(* IEC 61131-3 sources: NachHouse_TST/API/pilot_API_V10, 4 files *)

(* ---- 01_Nh_Api_STRUCT.st ---- *)
// NachHouse API PLC pilot V1.
// The public contract uses native PLCComS PUBLIC_API variables only.
// SK: Verejny kontrakt pouziva iba nativne PUBLIC_API premenne PLCComS.

VAR_GLOBAL CONSTANT
   NH_API_PROTOCOL_VERSION       : UINT := 1;            // Binary protocol version. SK: Verzia binarneho protokolu.
   NH_API_MAGIC                  : DWORD := 16#5041484E;  // ASCII NHAP bytes in little-endian order. SK: Bajty ASCII NHAP v little-endian poradi.
   NH_API_HEADER_SIZE            : UINT := 64;           // Fixed header size in bytes. SK: Pevna velkost hlavicky v bajtoch.
   NH_API_TX_WORD_COUNT          : UINT := 512;          // Number of DWORD words in the shared TX buffer. SK: Pocet DWORD slov spolocneho TX buffera.
   NH_API_RX_WORDS_PER_CLIENT    : UINT := 64;           // DWORD words in one client RX segment. SK: Pocet DWORD slov RX segmentu jedneho klienta.
   NH_API_RX_WORD_COUNT          : UINT := 256;          // Four RX segments of 64 DWORD each. SK: Styri RX segmenty po 64 DWORD.
   NH_API_MAX_CLIENTS            : USINT := 4;           // Maximum concurrently registered clients. SK: Najvacsi pocet sucasne registrovanych klientov.
   NH_API_MAX_ROOMS              : USINT := 40;          // Maximum number of pilot rooms. SK: Najvacsi pocet miestnosti pilotu.

   NH_API_CONFIG_RECORD_SIZE     : UINT := 138;          // Wire config record size. SK: Velkost wire config zaznamu.
   NH_API_STATE_RECORD_SIZE      : UINT := 22;           // Wire state record size including Twilight. SK: Velkost wire state zaznamu vratane Twilight.
   NH_API_CONFIG_DIFF_SIZE       : UINT := 143;          // Operation, RoomId and config record. SK: Operacia, RoomId a config zaznam.
   NH_API_STATE_DIFF_SIZE        : UINT := 27;           // Operation, RoomId and state record. SK: Operacia, RoomId a state zaznam.
   NH_API_CONFIG_PER_FRAME       : USINT := 14;          // Maximum config records in one TX frame. SK: Najviac config zaznamov v jednom TX ramci.
   NH_API_STATE_PER_FRAME        : USINT := 40;          // Maximum state records in one TX frame. SK: Najviac state zaznamov v jednom TX ramci.
   NH_API_CONFIG_DIFF_PER_FRAME  : USINT := 13;          // Maximum config changes in one TX frame. SK: Najviac config zmien v jednom TX ramci.
   NH_API_STATE_DIFF_PER_FRAME   : USINT := 40;          // Maximum state changes in one TX frame. SK: Najviac state zmien v jednom TX ramci.

   NH_API_TX_IDLE                : USINT := 0;            // TX buffer may be built. SK: TX buffer sa moze naplnit.
   NH_API_TX_BUILDING            : USINT := 1;            // PLC is building a TX frame. SK: PLC prave pripravuje TX ramec.
   NH_API_TX_READY               : USINT := 2;            // TX frame is stable and waiting for ACK. SK: TX ramec je stabilny a caka na ACK.

   NH_API_CLIENT_FREE            : USINT := 0;            // Client slot is free. SK: Klientsky slot je volny.
   NH_API_CLIENT_ACTIVE          : USINT := 1;            // Client slot has a valid lease. SK: Klientsky slot ma platny lease.

   NH_API_MSG_SNAPSHOT_REQUEST   : UINT := 1;             // RX full snapshot request. SK: RX poziadavka na kompletny snapshot.
   NH_API_MSG_ADD_ROOM           : UINT := 2;             // RX add-room request. SK: RX poziadavka na pridanie miestnosti.
   NH_API_MSG_DELETE_ROOM        : UINT := 3;             // RX delete-room request. SK: RX poziadavka na zmazanie miestnosti.
   NH_API_MSG_COPY_ROOM          : UINT := 4;             // RX copy-room request. SK: RX poziadavka na kopirovanie miestnosti.
   NH_API_MSG_SET_ROOM_CONFIG     : UINT := 5;             // RX room-config update request. SK: RX poziadavka na zmenu configu.
   NH_API_MSG_SET_ROOM_STATE      : UINT := 6;             // RX test room-state update request. SK: RX testovacia poziadavka na zmenu state.
   NH_API_MSG_CONFIG_SNAPSHOT    : UINT := 101;           // TX config snapshot part. SK: TX cast config snapshotu.
   NH_API_MSG_STATE_SNAPSHOT     : UINT := 102;           // TX state snapshot part. SK: TX cast state snapshotu.
   NH_API_MSG_CONFIG_DIFF        : UINT := 103;           // TX config diff. SK: TX config diff.
   NH_API_MSG_STATE_DIFF         : UINT := 104;           // TX state diff. SK: TX state diff.
   NH_API_MSG_SNAPSHOT_DONE      : UINT := 105;           // TX snapshot transaction completion. SK: TX ukoncenie snapshot transakcie.

   NH_API_SCHEMA_NONE            : UINT := 0;             // Message has no data record. SK: Sprava nema datovy zaznam.
   NH_API_SCHEMA_ROOM_CONFIG     : UINT := 1;             // Room configuration schema. SK: Schema konfiguracie miestnosti.
   NH_API_SCHEMA_ROOM_STATE      : UINT := 2;             // Room dynamic-state schema. SK: Schema dynamickeho stavu miestnosti.
   NH_API_SCHEMA_VERSION         : UINT := 1;             // Version of both room schemas. SK: Verzia oboch room schem.

   NH_API_CHANGE_UPSERT          : USINT := 1;            // Insert or complete record update. SK: Pridanie alebo uplna aktualizacia zaznamu.
   NH_API_CHANGE_DELETE          : USINT := 2;            // Record deletion. SK: Odstranenie zaznamu.

   NH_API_RESULT_NONE            : USINT := 0;            // No result is available yet. SK: Vysledok este neexistuje.
   NH_API_RESULT_OK              : USINT := 1;            // Request succeeded. SK: Poziadavka bola uspesna.
   NH_API_RESULT_BUSY            : USINT := 2;            // Another global transaction is active. SK: Ina globalna transakcia este bezi.
   NH_API_RESULT_BAD_FRAME       : USINT := 3;            // Header, size or CRC is invalid. SK: Hlavicka, velkost alebo CRC su neplatne.
   NH_API_RESULT_NOT_FOUND       : USINT := 4;            // Requested room does not exist. SK: Pozadovana miestnost neexistuje.
   NH_API_RESULT_NO_FREE_SLOT    : USINT := 5;            // No room or client slot is free. SK: Nie je volny room alebo client slot.
   NH_API_RESULT_ALREADY_EXISTS  : USINT := 6;            // RoomId already exists. SK: RoomId uz existuje.
   NH_API_RESULT_INVALID         : USINT := 7;            // Request payload is invalid. SK: Obsah poziadavky nie je platny.
   NH_API_RESULT_UNSUPPORTED     : USINT := 8;            // Message type is unsupported. SK: Typ spravy nie je podporovany.

   NH_API_TEST_NONE              : USINT := 0;            // WebMaker performs no action. SK: WebMaker nevykona ziadnu akciu.
   NH_API_TEST_SET_STATE         : USINT := 1;            // WebMaker changes room state. SK: WebMaker zmeni stav miestnosti.
   NH_API_TEST_ADD_ROOM          : USINT := 2;            // WebMaker adds a room. SK: WebMaker prida miestnost.
   NH_API_TEST_DELETE_ROOM       : USINT := 3;            // WebMaker deletes a room. SK: WebMaker zmaze miestnost.
   NH_API_TEST_COPY_ROOM         : USINT := 4;            // WebMaker copies a room. SK: WebMaker skopiruje miestnost.
   NH_API_TEST_SET_CONFIG        : USINT := 5;            // WebMaker changes room config. SK: WebMaker zmeni config miestnosti.
   NH_API_TEST_REQUEST_SNAPSHOT  : USINT := 6;            // WebMaker starts a broadcast snapshot. SK: WebMaker vyvola broadcast snapshot.
END_VAR

TYPE
   NH_ROOM_CONFIG : STRUCT // Static room configuration transferred in snapshots, diffs and commands. SK: Staticka konfiguracia miestnosti prenasana v snapshotoch, diffoch a prikazoch.
      Used           : BOOL;       // TRUE marks an occupied internal slot. SK: TRUE oznacuje obsadeny interny slot.
      RoomId         : UDINT;      // Stable unique room identifier. SK: Stabilny jedinecny identifikator miestnosti.
      Name           : STRING[64]; // UTF-8 room name, up to 64 bytes. SK: UTF-8 nazov miestnosti, najviac 64 bajtov.
      ProjectName    : STRING[64]; // UTF-8 project name, up to 64 bytes. SK: UTF-8 projektovy nazov, najviac 64 bajtov.
      IconId         : UINT;       // Client icon identifier. SK: Identifikator ikony klienta.
      SortDefault    : UINT;       // Default global order. SK: Predvolene globalne poradie.
   END_STRUCT

   NH_ROOM_STATE : STRUCT // Dynamic room state transferred in snapshots, diffs and commands. SK: Dynamicky stav miestnosti prenasany v snapshotoch, diffoch a prikazoch.
      RoomId         : UDINT;      // Stable ID matching the config record. SK: Stabilne ID zodpovedajuce config zaznamu.
      Temperature    : REAL;       // Temperature in degrees Celsius. SK: Teplota v stupnoch Celzia.
      Humidity       : REAL;       // Relative humidity in percent. SK: Relativna vlhkost v percentach.
      Presence       : BOOL;       // Presence flag. SK: Priznak pritomnosti.
      DayPhase       : UINT;       // Day-phase icon identifier. SK: Identifikator ikony dennej fazy.
      CategoryMask   : DWORD;      // Bit mask of active categories. SK: Bitova maska aktivnych kategorii.
      AlarmLevel     : USINT;      // Alarm level from 0 to 2. SK: Uroven alarmu 0 az 2.
      Online         : BOOL;       // Room data availability. SK: Dostupnost dat miestnosti.
      Twilight       : BOOL;       // Twilight state for the existing room browser. SK: Stav osvetlenia pre existujuci room browser.
   END_STRUCT

   NH_API_INFO : STRUCT // Global protocol, revision and shared TX-buffer handshake information. SK: Globalne informacie protokolu, revizii a handshake spolocneho TX buffera.
      ProtocolVersion : UINT;      // Wire protocol version. SK: Verzia wire protokolu.
      MaxRooms       : USINT;      // Number of available room slots. SK: Pocet dostupnych room slotov.
      MaxClients     : USINT;      // Number of client slots. SK: Pocet klientskych slotov.
      TxWordCount    : UINT;       // TX buffer size in DWORD words. SK: Velkost TX buffera v DWORD.
      RxWordsPerClient : UINT;     // One RX segment size in DWORD words. SK: Velkost jedneho RX segmentu v DWORD.
      ConfigRevision : UDINT;      // Current configuration revision. SK: Aktualna revizia konfiguracie.
      StateRevision  : UDINT;      // Current dynamic-state revision. SK: Aktualna revizia dynamickeho stavu.
      TxPublishedRevision : UDINT; // Commit identifier of the stable TX frame. SK: Commit identifikator stabilneho TX ramca.
      TxByteLength   : UINT;       // Number of valid TX frame bytes. SK: Pocet platnych bajtov TX ramca.
      TxState        : USINT;      // TX buffer state NH_API_TX_*. SK: Stav TX buffera NH_API_TX_*.
      TxRequiredAckMask : BYTE;    // Clients required to acknowledge the current frame. SK: Klienti, ktori musia potvrdit aktualny ramec.
      TxAckMask      : BYTE;       // Clients that already acknowledged the frame. SK: Klienti, ktori uz ramec potvrdili.
      ActiveClientMask : BYTE;     // Mask of valid client leases. SK: Maska platnych klientskych leases.
      LastError      : USINT;      // Last global diagnostic error. SK: Posledna globalna diagnosticka chyba.
   END_STRUCT

   NH_API_CLIENT_SLOT : STRUCT // Registration, liveness, RX commit and result state of one API client. SK: Registracia, zivotnost, RX commit a vysledkovy stav jedneho API klienta.
      RequestedClientId : UDINT;   // Random nonzero ID written by a registering client. SK: Nahodne nenulove ID zapisane klientom pri registracii.
      AssignedClientId : UDINT;    // ID accepted by the PLC for this slot. SK: ID potvrdene PLC pre tento slot.
      HeartbeatCounter : UDINT;    // Client periodically increments the liveness counter. SK: Klient periodicky zvysuje pocitadlo zivota.
      AckTxRevision : UDINT;       // Last TX frame whose CRC was verified. SK: Posledny TX ramec s overenym CRC.
      RxPublishedRevision : UDINT; // RX frame commit number written last by the client. SK: Commit cislo RX ramca zapisane klientom ako posledne.
      RxByteLength   : UINT;       // Valid byte count in the client RX segment. SK: Pocet platnych bajtov v klientovom RX segmente.
      State          : USINT;      // Registration state NH_API_CLIENT_*. SK: Stav registracie NH_API_CLIENT_*.
      ResultCode     : USINT;      // Result of the last accepted request. SK: Vysledok poslednej prijatej poziadavky.
      LastRequestId  : UDINT;      // RequestId belonging to ResultCode. SK: RequestId patriaci k ResultCode.
      ResultConfigRevision : UDINT;// Config revision after request execution. SK: Config revizia po vykonani poziadavky.
      ResultStateRevision : UDINT; // State revision after request execution. SK: State revizia po vykonani poziadavky.
   END_STRUCT

   NH_API_TEST_CONTROL : STRUCT // Direct WebMaker test interface used without a binary client. SK: Priame testovacie rozhranie WebMaker pouzivane bez binarneho klienta.
      Execute         : BOOL;       // WebMaker sets TRUE as the final commit step. SK: WebMaker nastavi TRUE ako posledny commit krok.
      Busy            : BOOL;       // PLC is processing the test action. SK: PLC prave spracovava testovaciu akciu.
      Finished        : BOOL;       // PLC completed the last test action. SK: PLC dokoncilo poslednu testovaciu akciu.
      Action          : USINT;      // Requested NH_API_TEST_* action. SK: Pozadovana akcia NH_API_TEST_*.
      ResultCode      : USINT;      // NH_API_RESULT_* outcome. SK: Vysledok NH_API_RESULT_*.
      RoomId          : UDINT;      // Target room ID. SK: Cielove ID miestnosti.
      SourceRoomId    : UDINT;      // Source ID for copying. SK: Zdrojove ID pri kopirovani.
      Name            : STRING[64]; // New name for add, copy or config update. SK: Novy nazov pre add, copy alebo set config.
      ProjectName     : STRING[64]; // New project name. SK: Novy projektovy nazov.
      IconId          : UINT;       // New room icon. SK: Nova ikona miestnosti.
      Temperature     : REAL;       // Test temperature. SK: Testovacia teplota.
      Humidity        : REAL;       // Test humidity. SK: Testovacia vlhkost.
      Presence        : BOOL;       // Test presence. SK: Testovacia pritomnost.
      DayPhase        : UINT;       // Test day phase. SK: Testovacia faza dna.
      CategoryMask    : DWORD;      // Test category mask. SK: Testovacia maska kategorii.
      AlarmLevel      : USINT;      // Test alarm level. SK: Testovacia uroven alarmu.
      Online          : BOOL;       // Test availability. SK: Testovacia dostupnost.
      Twilight        : BOOL;       // Test twilight state. SK: Testovaci twilight stav.
      ConfigRevision  : UDINT;      // Config revision after the action. SK: Config revizia po akcii.
      StateRevision   : UDINT;      // State revision after the action. SK: State revizia po akcii.
   END_STRUCT
END_TYPE

VAR_GLOBAL
   NH_API_CLIENT_TIMEOUT_MS      : UDINT := 500000;       // Time before an inactive client expires. SK: Cas do vyradenia neaktivneho klienta.

   NhApiInfo       {PUBLIC_API} : NH_API_INFO;                         // Global information and TX handshake. SK: Globalne informacie a TX handshake.
   NhApiClients    {PUBLIC_API} : ARRAY[0..3] OF NH_API_CLIENT_SLOT;   // Registry and handshake for four clients. SK: Registry a handshake styroch klientov.
   NhApiTxBuffer   {PUBLIC_API} : ARRAY[0..511] OF DWORD;              // Stable PLC-to-client message buffer. SK: Stabilny buffer sprav PLC smerom ku klientom.
   NhApiRxBuffer   {PUBLIC_API} : ARRAY[0..255] OF DWORD;              // Four separate client-to-PLC RX segments. SK: Styri oddelene klient-to-PLC RX segmenty.
   NhApiTest       {PUBLIC_API} : NH_API_TEST_CONTROL;                 // Direct WebMaker test control without a binary client. SK: Priamy WebMaker testovaci ovladac bez binarneho klienta.

   NhRoomsConfig                   : ARRAY[1..40] OF NH_ROOM_CONFIG;      // Authoritative PLC test configuration. SK: Autoritativna testovacia konfiguracia PLC.
   NhRoomsState                    : ARRAY[1..40] OF NH_ROOM_STATE;       // Authoritative PLC test state. SK: Autoritativny testovaci stav PLC.
END_VAR

VAR_GLOBAL
   NhApiInitialized                : BOOL;                                  // One-time initialization has completed. SK: Jednorazova inicializacia uz prebehla.
   NhConfigShadow                  : ARRAY[1..40] OF NH_ROOM_CONFIG;      // Last captured config used for diffing. SK: Posledny zachyteny config pre diff.
   NhStateShadow                   : ARRAY[1..40] OF NH_ROOM_STATE;       // Last captured state used for diffing. SK: Posledny zachyteny state pre diff.
   NhPendingConfig                 : ARRAY[1..40] OF NH_ROOM_CONFIG;      // Frozen config records of the current diff. SK: Zmrazene config zaznamy aktualneho diffu.
   NhPendingState                  : ARRAY[1..40] OF NH_ROOM_STATE;       // Frozen state records of the current diff. SK: Zmrazene state zaznamy aktualneho diffu.
   NhPendingOperation              : ARRAY[1..40] OF USINT;                 // Operations of the frozen diff. SK: Operacie zmrazeneho diffu.
   NhPendingRoomId                 : ARRAY[1..40] OF UDINT;                 // Room IDs of frozen diff items. SK: RoomId poloziek zmrazeneho diffu.
   NhPendingKind                   : UINT;                                  // Type of the pending config or state diff. SK: Typ rozpracovaneho config alebo state diffu.
   NhPendingCount                  : USINT;                                 // Number of pending diff items. SK: Pocet poloziek rozpracovaneho diffu.
   NhPendingNext                   : USINT;                                 // Index of the first item in the next frame. SK: Index prvej polozky dalsieho ramca.
   NhPendingPart                   : USINT;                                 // Number of the next diff part. SK: Cislo nasledujucej casti diffu.
   NhPendingParts                  : USINT;                                 // Total number of diff parts. SK: Celkovy pocet casti diffu.
   NhPendingFromRevision           : UDINT;                                // Starting domain revision of the diff. SK: Pociatocna domenova revizia diffu.
   NhPendingToRevision             : UDINT;                                // Ending domain revision of the diff. SK: Konecna domenova revizia diffu.

   NhSnapshotActive                : BOOL;                                  // A config-state-done sequence is active. SK: Prebieha sekvencia config-state-done.
   NhSnapshotTargetClientId        : UDINT;                                // Zero means broadcast, otherwise the target client. SK: Nula znamena broadcast, inak cielovy klient.
   NhSnapshotRequestId             : UDINT;                                // RequestId of the full snapshot. SK: RequestId kompletneho snapshotu.
   NhSnapshotStage                 : USINT;                                 // 1 config, 2 state, 3 done. SK: 1 config, 2 state, 3 done.
   NhSnapshotNext                  : USINT;                                 // First record index of the next part. SK: Index prveho zaznamu dalsej casti.
   NhSnapshotPart                  : USINT;                                 // Number of the next snapshot part. SK: Cislo dalsej casti snapshotu.
   NhSnapshotParts                 : USINT;                                 // Number of parts in the current snapshot section. SK: Pocet casti aktualnej snapshot sekcie.
   NhSnapshotConfig                : ARRAY[1..40] OF NH_ROOM_CONFIG;      // Frozen config portion of the snapshot. SK: Zmrazena config cast snapshotu.
   NhSnapshotState                 : ARRAY[1..40] OF NH_ROOM_STATE;       // Frozen state portion of the snapshot. SK: Zmrazena state cast snapshotu.
   NhSnapshotCount                 : USINT;                                 // Number of valid snapshot rooms. SK: Pocet platnych miestnosti snapshotu.

   NhClientLastHeartbeat           : ARRAY[0..3] OF UDINT;                  // Last processed heartbeat values. SK: Posledne spracovane heartbeat hodnoty.
   NhClientLastAck                 : ARRAY[0..3] OF UDINT;                  // Last processed ACK values. SK: Posledne spracovane ACK hodnoty.
   NhClientLastRx                  : ARRAY[0..3] OF UDINT;                  // Last processed RX commit values. SK: Posledne spracovane RX commit hodnoty.
   NhClientLastActivityMs          : ARRAY[0..3] OF UDINT;                  // System time of the last activity. SK: Systemovy cas poslednej aktivity.
END_VAR

(* ---- 02_Nh_Api_UTILS.st ---- *)
// Wire-format helpers have no hidden state. SK: Pomocne funkcie wire formatu su bez skryteho stavu.

FUNCTION NhApiNextRevision : UDINT
   // Returns the next nonzero revision. SK: Vrati nasledujucu nenulovu reviziu.
   VAR_INPUT
      Current : UDINT; // Current revision. SK: Aktualna revizia.
   END_VAR
   NhApiNextRevision := Current + 1;
   IF NhApiNextRevision = 0 THEN
      NhApiNextRevision := 1;
   END_IF;
END_FUNCTION

FUNCTION NhApiSystemTimeMs : UDINT
   // Returns the PLC system time in milliseconds. SK: Vrati systemovy cas PLC v milisekundach.
   VAR_EXTERNAL
      AT %SL52 : DWORD; // Absolute PLC system-time register. SK: Absolutny systemovy register casu PLC.
   END_VAR
   NhApiSystemTimeMs := DWORD_TO_UDINT(%SL52);
END_FUNCTION

FUNCTION NhApiWriteByte : BOOL
   // Writes one byte at the specified buffer offset. SK: Zapise jeden bajt na zadany offset buffera.
   VAR_INPUT
      Buffer : PTR_TO BYTE; // Start of the destination buffer. SK: Zaciatok cieloveho buffera.
      Offset : UINT;        // Zero-based byte offset. SK: Nulovy byte offset.
      Value  : BYTE;        // Value to write. SK: Zapisovana hodnota.
   END_VAR
   VAR
      Position : PTR_TO BYTE; // Pointer advanced to the target byte. SK: Pointer posunuty na cielovy bajt.
   END_VAR
   Position := Buffer + UINT_TO_UDINT(Offset);
   Position^ := Value;
   NhApiWriteByte := TRUE;
END_FUNCTION

FUNCTION NhApiReadByte : BYTE
   // Reads one byte from the specified buffer offset. SK: Precita jeden bajt zo zadaneho offsetu buffera.
   VAR_INPUT
      Buffer : PTR_TO BYTE; // Start of the source buffer. SK: Zaciatok zdrojoveho buffera.
      Offset : UINT;        // Zero-based byte offset. SK: Nulovy byte offset.
   END_VAR
   VAR
      Position : PTR_TO BYTE; // Pointer advanced to the source byte. SK: Pointer posunuty na zdrojovy bajt.
   END_VAR
   Position := Buffer + UINT_TO_UDINT(Offset);
   NhApiReadByte := Position^;
END_FUNCTION

FUNCTION NhApiWriteU16 : BOOL
   // Writes a 16-bit value in little-endian format. SK: Zapise 16-bitovu hodnotu vo formate little-endian.
   VAR_INPUT
      Buffer : PTR_TO BYTE; // Destination byte buffer. SK: Cielovy byte buffer.
      Offset : UINT;        // Zero-based byte offset. SK: Nulovy byte offset.
      Value  : UINT;        // Value written little-endian. SK: Hodnota zapisovana little-endian.
   END_VAR
   NhApiWriteByte(Buffer := Buffer, Offset := Offset, Value := WORD_TO_BYTE(UINT_TO_WORD(Value) AND 16#00FF));
   NhApiWriteByte(Buffer := Buffer, Offset := Offset + 1, Value := WORD_TO_BYTE(SHR(UINT_TO_WORD(Value), 8)));
   NhApiWriteU16 := TRUE;
END_FUNCTION

FUNCTION NhApiWriteU32 : BOOL
   // Writes a 32-bit value in little-endian format. SK: Zapise 32-bitovu hodnotu vo formate little-endian.
   VAR_INPUT
      Buffer : PTR_TO BYTE; // Destination byte buffer. SK: Cielovy byte buffer.
      Offset : UINT;        // Zero-based byte offset. SK: Nulovy byte offset.
      Value  : UDINT;       // Value written little-endian. SK: Hodnota zapisovana little-endian.
   END_VAR
   VAR
      Raw : DWORD;          // Bit image of the value. SK: Bitovy obraz hodnoty.
   END_VAR
   Raw := UDINT_TO_DWORD(Value);
   NhApiWriteByte(Buffer := Buffer, Offset := Offset, Value := DWORD_TO_BYTE(Raw AND 16#000000FF));
   NhApiWriteByte(Buffer := Buffer, Offset := Offset + 1, Value := DWORD_TO_BYTE(SHR(Raw, 8) AND 16#000000FF));
   NhApiWriteByte(Buffer := Buffer, Offset := Offset + 2, Value := DWORD_TO_BYTE(SHR(Raw, 16) AND 16#000000FF));
   NhApiWriteByte(Buffer := Buffer, Offset := Offset + 3, Value := DWORD_TO_BYTE(SHR(Raw, 24) AND 16#000000FF));
   NhApiWriteU32 := TRUE;
END_FUNCTION

FUNCTION NhApiReadU16 : UINT
   // Reads a 16-bit value in little-endian format. SK: Precita 16-bitovu hodnotu vo formate little-endian.
   VAR_INPUT
      Buffer : PTR_TO BYTE; // Source byte buffer. SK: Zdrojovy byte buffer.
      Offset : UINT;        // Zero-based byte offset. SK: Nulovy byte offset.
   END_VAR
   NhApiReadU16 := WORD_TO_UINT(BYTE_TO_WORD(NhApiReadByte(Buffer := Buffer, Offset := Offset)) OR
      SHL(BYTE_TO_WORD(NhApiReadByte(Buffer := Buffer, Offset := Offset + 1)), 8));
END_FUNCTION

FUNCTION NhApiReadU32 : UDINT
   // Reads a 32-bit value in little-endian format. SK: Precita 32-bitovu hodnotu vo formate little-endian.
   VAR_INPUT
      Buffer : PTR_TO BYTE; // Source byte buffer. SK: Zdrojovy byte buffer.
      Offset : UINT;        // Zero-based byte offset. SK: Nulovy byte offset.
   END_VAR
   VAR
      Raw : DWORD;          // Reassembled little-endian value. SK: Zlozena little-endian hodnota.
   END_VAR
   Raw := BYTE_TO_DWORD(NhApiReadByte(Buffer := Buffer, Offset := Offset));
   Raw := Raw OR SHL(BYTE_TO_DWORD(NhApiReadByte(Buffer := Buffer, Offset := Offset + 1)), 8);
   Raw := Raw OR SHL(BYTE_TO_DWORD(NhApiReadByte(Buffer := Buffer, Offset := Offset + 2)), 16);
   Raw := Raw OR SHL(BYTE_TO_DWORD(NhApiReadByte(Buffer := Buffer, Offset := Offset + 3)), 24);
   NhApiReadU32 := DWORD_TO_UDINT(Raw);
END_FUNCTION

FUNCTION NhApiWriteReal : BOOL
   // Writes a REAL using its 32-bit image. SK: Zapise REAL pomocou jeho 32-bitoveho obrazu.
   VAR_INPUT
      Buffer : PTR_TO BYTE; // Destination byte buffer. SK: Cielovy byte buffer.
      Offset : UINT;        // Zero-based byte offset. SK: Nulovy byte offset.
      Value  : REAL;        // IEC REAL written by bit image. SK: IEC REAL zapisany bitovo.
   END_VAR
   VAR
      RawPtr : PTR_TO DWORD;// Pointer to the REAL bit image. SK: Pointer na bitovy obraz REAL.
   END_VAR
   RawPtr := ADR(Value);
   NhApiWriteU32(Buffer := Buffer, Offset := Offset, Value := DWORD_TO_UDINT(RawPtr^));
   NhApiWriteReal := TRUE;
END_FUNCTION

FUNCTION NhApiReadReal : REAL
   // Reads a REAL from its 32-bit image. SK: Precita REAL z jeho 32-bitoveho obrazu.
   VAR_INPUT
      Buffer : PTR_TO BYTE; // Source byte buffer. SK: Zdrojovy byte buffer.
      Offset : UINT;        // Zero-based byte offset. SK: Nulovy byte offset.
   END_VAR
   VAR
      ResultPtr : PTR_TO DWORD; // Pointer to the result bit image. SK: Pointer na bitovy obraz vysledku.
   END_VAR
   ResultPtr := ADR(NhApiReadReal);
   ResultPtr^ := UDINT_TO_DWORD(NhApiReadU32(Buffer := Buffer, Offset := Offset));
END_FUNCTION

FUNCTION NhApiFrameCrc32 : DWORD
   // Calculates CRC32 of the valid API frame. SK: Vypocita CRC32 platnej casti API ramca.
   VAR_INPUT
      Buffer : PTR_TO BYTE; // Start of the complete frame. SK: Zaciatok celeho ramca.
      Length : UINT;        // Header plus payload. SK: Hlavicka plus payload.
   END_VAR
   VAR
      Crc       : DWORD;    // Running CRC32 value. SK: PriebeznA CRC32 hodnota.
      Current   : BYTE;     // Current byte; CRC field is treated as zero. SK: Aktualny bajt; CRC pole sa pocita ako nula.
      Index     : UINT;     // Byte index. SK: Index bajtu.
      BitIndex  : USINT;    // Bit index. SK: Index bitu.
   END_VAR
   Crc := 16#FFFFFFFF;
   IF Length > 0 THEN
      FOR Index := 0 TO Length - 1 DO
         IF (Index >= 60) AND (Index <= 63) THEN
            Current := 0;
         ELSE
            Current := NhApiReadByte(Buffer := Buffer, Offset := Index);
         END_IF;
         Crc := Crc XOR BYTE_TO_DWORD(Current);
         FOR BitIndex := 0 TO 7 DO
            IF (Crc AND 16#00000001) <> 0 THEN
               Crc := SHR(Crc, 1) XOR 16#EDB88320;
            ELSE
               Crc := SHR(Crc, 1);
            END_IF;
         END_FOR;
      END_FOR;
   END_IF;
   NhApiFrameCrc32 := NOT Crc;
END_FUNCTION

FUNCTION NhApiClearBuffer : BOOL
   // Clears the specified number of buffer bytes. SK: Vynuluje zadany pocet bajtov buffera.
   VAR_INPUT
      Buffer : PTR_TO BYTE; // Buffer to clear. SK: Buffer urceny na vynulovanie.
      Length : UINT;        // Number of bytes. SK: Pocet bajtov.
   END_VAR
   VAR
      Index : UINT;         // Index of the cleared byte. SK: Index nulovaneho bajtu.
   END_VAR
   IF Length > 0 THEN
      FOR Index := 0 TO Length - 1 DO
         NhApiWriteByte(Buffer := Buffer, Offset := Index, Value := 0);
      END_FOR;
   END_IF;
   NhApiClearBuffer := TRUE;
END_FUNCTION

FUNCTION NhApiConfigEqual : BOOL
   // Compares two room configuration records. SK: Porovna dva konfiguracne zaznamy miestnosti.
   VAR_INPUT
      A : NH_ROOM_CONFIG; // First config record. SK: Prvy config zaznam.
      B : NH_ROOM_CONFIG; // Second config record. SK: Druhy config zaznam.
   END_VAR
   NhApiConfigEqual := (A.Used = B.Used) AND (A.RoomId = B.RoomId) AND (A.Name = B.Name) AND
      (A.ProjectName = B.ProjectName) AND (A.IconId = B.IconId) AND (A.SortDefault = B.SortDefault);
END_FUNCTION

FUNCTION NhApiStateEqual : BOOL
   // Compares two dynamic room-state records. SK: Porovna dva dynamicke stavove zaznamy miestnosti.
   VAR_INPUT
      A : NH_ROOM_STATE;  // First state record. SK: Prvy state zaznam.
      B : NH_ROOM_STATE;  // Second state record. SK: Druhy state zaznam.
   END_VAR
   NhApiStateEqual := (A.RoomId = B.RoomId) AND (A.Temperature = B.Temperature) AND
      (A.Humidity = B.Humidity) AND (A.Presence = B.Presence) AND (A.DayPhase = B.DayPhase) AND
      (A.CategoryMask = B.CategoryMask) AND (A.AlarmLevel = B.AlarmLevel) AND
      (A.Online = B.Online) AND (A.Twilight = B.Twilight);
END_FUNCTION

FUNCTION NhApiFindRoom : USINT
   // Finds a room slot by its stable ID. SK: Najde interny slot miestnosti podla stabilneho ID.
   VAR_INPUT
      RoomId : UDINT;       // Stable ID to find. SK: Hladane stabilne ID.
   END_VAR
   VAR
      Index : USINT;        // Index of the scanned slot. SK: Index prehladavaneho slotu.
   END_VAR
   NhApiFindRoom := 0;
   FOR Index := 1 TO NH_API_MAX_ROOMS DO
      IF NhRoomsConfig[Index].Used AND (NhRoomsConfig[Index].RoomId = RoomId) THEN
         NhApiFindRoom := Index;
         RETURN;
      END_IF;
   END_FOR;
END_FUNCTION

FUNCTION NhApiFindFreeRoom : USINT
   // Finds the first free internal room slot. SK: Najde prvy volny interny slot miestnosti.
   VAR
      Index : USINT;        // Index of the scanned slot. SK: Index prehladavaneho slotu.
   END_VAR
   NhApiFindFreeRoom := 0;
   FOR Index := 1 TO NH_API_MAX_ROOMS DO
      IF NOT NhRoomsConfig[Index].Used THEN
         NhApiFindFreeRoom := Index;
         RETURN;
      END_IF;
   END_FOR;
END_FUNCTION

FUNCTION NhApiWriteText64 : BOOL
   // Writes text into a fixed 65-byte wire field. SK: Zapise text do pevneho 65-bajtoveho wire pola.
   VAR_INPUT
      Buffer : PTR_TO BYTE; // Destination wire buffer. SK: Cielovy wire buffer.
      Offset : UINT;        // Offset of length and 64 text bytes. SK: Offset dlzky a 64 bajtov textu.
      Value  : STRING[64];  // UTF-8 bytes stored in the PLC STRING. SK: UTF-8 bajty ulozene v PLC STRING.
   END_VAR
   VAR
      Source : PTR_TO BYTE; // First PLC STRING byte. SK: Prvy bajt PLC STRING.
      Index  : USINT;       // Text byte index. SK: Index textoveho bajtu.
      Count  : USINT;       // Number of actual bytes. SK: Pocet skutocnych bajtov.
   END_VAR
   Count := INT_TO_USINT(LEN(Value));
   IF Count > 64 THEN
      Count := 64;
   END_IF;
   NhApiWriteByte(Buffer := Buffer, Offset := Offset, Value := USINT_TO_BYTE(Count));
   Source := ADR(Value);
   FOR Index := 0 TO 63 DO
      IF Index < Count THEN
         NhApiWriteByte(Buffer := Buffer, Offset := Offset + 1 + USINT_TO_UINT(Index),
            Value := NhApiReadByte(Buffer := Source, Offset := USINT_TO_UINT(Index)));
      ELSE
         NhApiWriteByte(Buffer := Buffer, Offset := Offset + 1 + USINT_TO_UINT(Index), Value := 0);
      END_IF;
   END_FOR;
   NhApiWriteText64 := TRUE;
END_FUNCTION

FUNCTION NhApiReadText64 : STRING[64]
   // Reads text from a fixed 65-byte wire field. SK: Precita text z pevneho 65-bajtoveho wire pola.
   VAR_INPUT
      Buffer : PTR_TO BYTE; // Source wire buffer. SK: Zdrojovy wire buffer.
      Offset : UINT;        // Offset of length and 64 text bytes. SK: Offset dlzky a 64 bajtov textu.
   END_VAR
   VAR
      Destination : PTR_TO BYTE; // First byte of the result PLC STRING. SK: Prvy bajt vysledneho PLC STRING.
      Index       : USINT;       // Text byte index. SK: Index textoveho bajtu.
      Count       : USINT;       // Declared byte count. SK: Deklarovany pocet bajtov.
   END_VAR
   Count := BYTE_TO_USINT(NhApiReadByte(Buffer := Buffer, Offset := Offset));
   IF Count > 64 THEN
      Count := 64;
   END_IF;
   Destination := ADR(NhApiReadText64);
   FOR Index := 0 TO 63 DO
      IF Index < Count THEN
         NhApiWriteByte(Buffer := Destination, Offset := USINT_TO_UINT(Index),
            Value := NhApiReadByte(Buffer := Buffer, Offset := Offset + 1 + USINT_TO_UINT(Index)));
      ELSE
         NhApiWriteByte(Buffer := Destination, Offset := USINT_TO_UINT(Index), Value := 0);
      END_IF;
   END_FOR;
END_FUNCTION

FUNCTION NhApiWriteConfigRecord : BOOL
   // Serializes a room configuration record. SK: Serializuje konfiguracny zaznam miestnosti.
   VAR_INPUT
      Buffer : PTR_TO BYTE;       // Destination wire buffer. SK: Cielovy wire buffer.
      Offset : UINT;              // Record start offset. SK: Offset zaciatku zaznamu.
      Record : NH_ROOM_CONFIG;  // Config record to serialize. SK: Config zaznam na serializaciu.
   END_VAR
   NhApiWriteU32(Buffer := Buffer, Offset := Offset, Value := Record.RoomId);
   NhApiWriteU16(Buffer := Buffer, Offset := Offset + 4, Value := Record.IconId);
   NhApiWriteU16(Buffer := Buffer, Offset := Offset + 6, Value := Record.SortDefault);
   NhApiWriteText64(Buffer := Buffer, Offset := Offset + 8, Value := Record.Name);
   NhApiWriteText64(Buffer := Buffer, Offset := Offset + 73, Value := Record.ProjectName);
   NhApiWriteConfigRecord := TRUE;
END_FUNCTION

FUNCTION NhApiReadConfigRecord : BOOL
   // Deserializes a room configuration record. SK: Deserializuje konfiguracny zaznam miestnosti.
   VAR_INPUT
      Buffer : PTR_TO BYTE;       // Source wire buffer. SK: Zdrojovy wire buffer.
      Offset : UINT;              // Record start offset. SK: Offset zaciatku zaznamu.
   END_VAR
   VAR_IN_OUT
      Record : NH_ROOM_CONFIG;  // Decoded config record. SK: Dekodovany config zaznam.
   END_VAR
   Record.Used := TRUE;
   Record.RoomId := NhApiReadU32(Buffer := Buffer, Offset := Offset);
   Record.IconId := NhApiReadU16(Buffer := Buffer, Offset := Offset + 4);
   Record.SortDefault := NhApiReadU16(Buffer := Buffer, Offset := Offset + 6);
   Record.Name := NhApiReadText64(Buffer := Buffer, Offset := Offset + 8);
   Record.ProjectName := NhApiReadText64(Buffer := Buffer, Offset := Offset + 73);
   NhApiReadConfigRecord := TRUE;
END_FUNCTION

FUNCTION NhApiWriteStateRecord : BOOL
   // Serializes a dynamic room-state record. SK: Serializuje dynamicky stavovy zaznam miestnosti.
   VAR_INPUT
      Buffer : PTR_TO BYTE;       // Destination wire buffer. SK: Cielovy wire buffer.
      Offset : UINT;              // Record start offset. SK: Offset zaciatku zaznamu.
      Record : NH_ROOM_STATE;   // State record to serialize. SK: State zaznam na serializaciu.
   END_VAR
   NhApiWriteU32(Buffer := Buffer, Offset := Offset, Value := Record.RoomId);
   NhApiWriteReal(Buffer := Buffer, Offset := Offset + 4, Value := Record.Temperature);
   NhApiWriteReal(Buffer := Buffer, Offset := Offset + 8, Value := Record.Humidity);
   NhApiWriteByte(Buffer := Buffer, Offset := Offset + 12, Value := BOOL_TO_BYTE(Record.Presence));
   NhApiWriteU16(Buffer := Buffer, Offset := Offset + 13, Value := Record.DayPhase);
   NhApiWriteU32(Buffer := Buffer, Offset := Offset + 15, Value := DWORD_TO_UDINT(Record.CategoryMask));
   NhApiWriteByte(Buffer := Buffer, Offset := Offset + 19, Value := USINT_TO_BYTE(Record.AlarmLevel));
   NhApiWriteByte(Buffer := Buffer, Offset := Offset + 20, Value := BOOL_TO_BYTE(Record.Online));
   NhApiWriteByte(Buffer := Buffer, Offset := Offset + 21, Value := BOOL_TO_BYTE(Record.Twilight));
   NhApiWriteStateRecord := TRUE;
END_FUNCTION

FUNCTION NhApiReadStateRecord : BOOL
   // Deserializes a dynamic room-state record. SK: Deserializuje dynamicky stavovy zaznam miestnosti.
   VAR_INPUT
      Buffer : PTR_TO BYTE;       // Source wire buffer. SK: Zdrojovy wire buffer.
      Offset : UINT;              // Record start offset. SK: Offset zaciatku zaznamu.
   END_VAR
   VAR_IN_OUT
      Record : NH_ROOM_STATE;   // Decoded state record. SK: Dekodovany state zaznam.
   END_VAR
   Record.RoomId := NhApiReadU32(Buffer := Buffer, Offset := Offset);
   Record.Temperature := NhApiReadReal(Buffer := Buffer, Offset := Offset + 4);
   Record.Humidity := NhApiReadReal(Buffer := Buffer, Offset := Offset + 8);
   Record.Presence := NhApiReadByte(Buffer := Buffer, Offset := Offset + 12) <> 0;
   Record.DayPhase := NhApiReadU16(Buffer := Buffer, Offset := Offset + 13);
   Record.CategoryMask := UDINT_TO_DWORD(NhApiReadU32(Buffer := Buffer, Offset := Offset + 15));
   Record.AlarmLevel := BYTE_TO_USINT(NhApiReadByte(Buffer := Buffer, Offset := Offset + 19));
   Record.Online := NhApiReadByte(Buffer := Buffer, Offset := Offset + 20) <> 0;
   Record.Twilight := NhApiReadByte(Buffer := Buffer, Offset := Offset + 21) <> 0;
   NhApiReadStateRecord := TRUE;
END_FUNCTION

(* ---- 03_Nh_Api_ENGINE.st ---- *)
// State machine, application operations and frame publishing. SK: Stavovy automat, aplikacne operacie a publikovanie ramcov.

FUNCTION NhApiClearRoom : BOOL
   // Clears the configuration and state of one room slot. SK: Vynuluje konfiguraciu a stav jedneho room slotu.
   VAR_INPUT
      Index : USINT; // Internal room slot 1..40. SK: Interny room slot 1..40.
   END_VAR
   NhRoomsConfig[Index].Used := FALSE;
   NhRoomsConfig[Index].RoomId := 0;
   NhRoomsConfig[Index].Name := '';
   NhRoomsConfig[Index].ProjectName := '';
   NhRoomsConfig[Index].IconId := 0;
   NhRoomsConfig[Index].SortDefault := 0;
   NhRoomsState[Index].RoomId := 0;
   NhRoomsState[Index].Temperature := 0.0;
   NhRoomsState[Index].Humidity := 0.0;
   NhRoomsState[Index].Presence := FALSE;
   NhRoomsState[Index].DayPhase := 140;
   NhRoomsState[Index].CategoryMask := 0;
   NhRoomsState[Index].AlarmLevel := 0;
   NhRoomsState[Index].Online := FALSE;
   NhRoomsState[Index].Twilight := FALSE;
   NhApiClearRoom := TRUE;
END_FUNCTION

FUNCTION NhApiInitialize : BOOL
   // Initializes API data, buffers, and state once. SK: Jednorazovo inicializuje data, buffery a stav API.
   VAR
      Index : USINT; // Initialization index. SK: Inicializacny index.
   END_VAR
   NhApiInitialize := NhApiInitialized;
   IF NhApiInitialized THEN
      RETURN;
   END_IF;

   NhApiClearBuffer(Buffer := ADR(NhApiTxBuffer), Length := 2048);
   NhApiClearBuffer(Buffer := ADR(NhApiRxBuffer), Length := 1024);
   FOR Index := 1 TO NH_API_MAX_ROOMS DO
      NhApiClearRoom(Index := Index);
   END_FOR;

   // Thirty deterministic ASCII names are also valid UTF-8. SK: Tridsat deterministickych ASCII nazvov je sucasne platne UTF-8.
   FOR Index := 1 TO 30 DO
      NhRoomsConfig[Index].Used := TRUE;
      NhRoomsConfig[Index].RoomId := USINT_TO_UDINT(Index);
      NhRoomsConfig[Index].ProjectName := 'TEST';
      NhRoomsConfig[Index].IconId := SEL(Index >= 26, 16, 19);
      NhRoomsConfig[Index].SortDefault := USINT_TO_UINT(Index);
      CASE Index OF
         1: NhRoomsConfig[Index].Name := 'Hall 1'; NhRoomsConfig[Index].ProjectName := '1.08';
         2: NhRoomsConfig[Index].Name := 'Kitchen'; NhRoomsConfig[Index].ProjectName := '1.07';
         3: NhRoomsConfig[Index].Name := 'Corridor 1'; NhRoomsConfig[Index].ProjectName := '1.04';
         4: NhRoomsConfig[Index].Name := 'Bathroom 1'; NhRoomsConfig[Index].ProjectName := '1.06';
         5: NhRoomsConfig[Index].Name := 'WC'; NhRoomsConfig[Index].ProjectName := '1.05';
         6: NhRoomsConfig[Index].Name := 'Bedroom'; NhRoomsConfig[Index].ProjectName := '1.09';
         7: NhRoomsConfig[Index].Name := 'Boiler'; NhRoomsConfig[Index].ProjectName := '1.03';
         8: NhRoomsConfig[Index].Name := 'Living room'; NhRoomsConfig[Index].ProjectName := '1.01';
         9: NhRoomsConfig[Index].Name := 'Corridor 1F'; NhRoomsConfig[Index].ProjectName := '1.02';
         10: NhRoomsConfig[Index].Name := 'Room 2.07'; NhRoomsConfig[Index].ProjectName := '2.07';
         11: NhRoomsConfig[Index].Name := 'Kitchen 2F'; NhRoomsConfig[Index].ProjectName := '2.03';
         12: NhRoomsConfig[Index].Name := 'Room 2.06'; NhRoomsConfig[Index].ProjectName := '2.06';
         13: NhRoomsConfig[Index].Name := 'Bathroom 2F'; NhRoomsConfig[Index].ProjectName := '2.05';
         14: NhRoomsConfig[Index].Name := 'Entrance hall'; NhRoomsConfig[Index].ProjectName := '0.01';
         15: NhRoomsConfig[Index].Name := 'Garage'; NhRoomsConfig[Index].ProjectName := '0.02';
         16: NhRoomsConfig[Index].Name := 'Storage'; NhRoomsConfig[Index].ProjectName := '0.03';
         17: NhRoomsConfig[Index].Name := 'Basement corridor'; NhRoomsConfig[Index].ProjectName := '0.04';
         18: NhRoomsConfig[Index].Name := 'Office'; NhRoomsConfig[Index].ProjectName := '1.10';
         19: NhRoomsConfig[Index].Name := 'Wardrobe'; NhRoomsConfig[Index].ProjectName := '1.11';
         20: NhRoomsConfig[Index].Name := 'Fitness'; NhRoomsConfig[Index].ProjectName := '0.06';
         21: NhRoomsConfig[Index].Name := 'Technical'; NhRoomsConfig[Index].ProjectName := '0.07';
         22: NhRoomsConfig[Index].Name := 'Wine room'; NhRoomsConfig[Index].ProjectName := '0.08';
         23: NhRoomsConfig[Index].Name := 'Guest room'; NhRoomsConfig[Index].ProjectName := '2.01';
         24: NhRoomsConfig[Index].Name := 'Children 1'; NhRoomsConfig[Index].ProjectName := '2.02';
         25: NhRoomsConfig[Index].Name := 'Children 2'; NhRoomsConfig[Index].ProjectName := '2.04';
         26: NhRoomsConfig[Index].Name := 'Terrace'; NhRoomsConfig[Index].ProjectName := 'E.01';
         27: NhRoomsConfig[Index].Name := 'Gazebo'; NhRoomsConfig[Index].ProjectName := 'E.02';
         28: NhRoomsConfig[Index].Name := 'Pool'; NhRoomsConfig[Index].ProjectName := 'E.03';
         29: NhRoomsConfig[Index].Name := 'Garden'; NhRoomsConfig[Index].ProjectName := 'E.04';
         30: NhRoomsConfig[Index].Name := 'Sauna'; NhRoomsConfig[Index].ProjectName := '0.09';
      END_CASE;
      NhRoomsState[Index].RoomId := USINT_TO_UDINT(Index);
      NhRoomsState[Index].Temperature := 20.0 + USINT_TO_REAL(Index) * 0.1;
      NhRoomsState[Index].Humidity := 40.0 + USINT_TO_REAL(Index MOD 15);
      NhRoomsState[Index].Presence := (Index MOD 4) = 0;
      CASE Index MOD 4 OF
         0: NhRoomsState[Index].DayPhase := 140;
         1: NhRoomsState[Index].DayPhase := 142;
         2: NhRoomsState[Index].DayPhase := 144;
         3: NhRoomsState[Index].DayPhase := 146;
      END_CASE;
      NhRoomsState[Index].CategoryMask := USINT_TO_DWORD(Index MOD 8);
      NhRoomsState[Index].AlarmLevel := 0;
      NhRoomsState[Index].Online := (Index MOD 3) <> 0;
      NhRoomsState[Index].Twilight := (Index MOD 3) <> 1;
      NhConfigShadow[Index] := NhRoomsConfig[Index];
      NhStateShadow[Index] := NhRoomsState[Index];
   END_FOR;
   FOR Index := 31 TO NH_API_MAX_ROOMS DO
      NhConfigShadow[Index] := NhRoomsConfig[Index];
      NhStateShadow[Index] := NhRoomsState[Index];
   END_FOR;

   NhApiInfo.ProtocolVersion := NH_API_PROTOCOL_VERSION;
   NhApiInfo.MaxRooms := NH_API_MAX_ROOMS;
   NhApiInfo.MaxClients := NH_API_MAX_CLIENTS;
   NhApiInfo.TxWordCount := NH_API_TX_WORD_COUNT;
   NhApiInfo.RxWordsPerClient := NH_API_RX_WORDS_PER_CLIENT;
   NhApiInfo.ConfigRevision := 1;
   NhApiInfo.StateRevision := 1;
   NhApiInfo.TxPublishedRevision := 0;
   NhApiInfo.TxByteLength := 0;
   NhApiInfo.TxState := NH_API_TX_IDLE;
   NhApiInfo.TxRequiredAckMask := 0;
   NhApiInfo.TxAckMask := 0;
   NhApiInfo.ActiveClientMask := 0;
   NhApiInfo.LastError := NH_API_RESULT_NONE;
   FOR Index := 0 TO 3 DO
      NhApiClients[Index].RequestedClientId := 0;
      NhApiClients[Index].AssignedClientId := 0;
      NhApiClients[Index].HeartbeatCounter := 0;
      NhApiClients[Index].AckTxRevision := 0;
      NhApiClients[Index].RxPublishedRevision := 0;
      NhApiClients[Index].RxByteLength := 0;
      NhApiClients[Index].State := NH_API_CLIENT_FREE;
      NhApiClients[Index].ResultCode := NH_API_RESULT_NONE;
      NhApiClients[Index].LastRequestId := 0;
      NhApiClients[Index].ResultConfigRevision := 1;
      NhApiClients[Index].ResultStateRevision := 1;
      NhClientLastActivityMs[Index] := NhApiSystemTimeMs();
   END_FOR;
   NhApiTest.Execute := FALSE;
   NhApiTest.Busy := FALSE;
   NhApiTest.Finished := FALSE;
   NhApiTest.ResultCode := NH_API_RESULT_NONE;
   NhPendingKind := 0;
   NhSnapshotActive := FALSE;
   NhApiInitialized := TRUE;
   NhApiInitialize := TRUE;
END_FUNCTION

FUNCTION NhApiBeginFrame : BOOL
   // Prepares a new TX frame header and clears the TX buffer. SK: Pripravi hlavicku noveho TX ramca a vycisti TX buffer.
   VAR_INPUT
      MessageType : UINT;   // TX message type. SK: Typ TX spravy.
      SchemaId : UINT;      // Record schema identifier. SK: Identifikator record schemy.
      TargetClientId : UDINT;// Zero for broadcast. SK: Nula pre broadcast.
      RequestId : UDINT;    // Original RequestId or zero. SK: Povodny RequestId alebo nula.
      FromRevision : UDINT; // Previous domain revision. SK: Predchadzajuca domenova revizia.
      ToRevision : UDINT;   // New domain revision. SK: Nova domenova revizia.
      RecordCount : UINT;   // Number of records in payload. SK: Pocet zaznamov v payload.
      RecordSize : UINT;    // Fixed size of one record. SK: Pevna velkost jedneho zaznamu.
      PartIndex : UINT;     // One-based part number. SK: Jednotkove cislo casti.
      PartCount : UINT;     // Total number of parts. SK: Celkovy pocet casti.
   END_VAR
   VAR
      Buffer : PTR_TO BYTE; // Byte view of the TX DWORD array. SK: Byte pohlad na TX DWORD pole.
      PayloadSize : UDINT;  // Calculated payload size. SK: Vypocitana velkost payloadu.
      TotalSize : UDINT;    // Header plus payload. SK: Hlavicka plus payload.
      FrameRevision : UDINT;// New frame transport revision. SK: Nova transportna revizia ramca.
   END_VAR
   Buffer := ADR(NhApiTxBuffer);
   NhApiInfo.TxState := NH_API_TX_BUILDING;
   NhApiClearBuffer(Buffer := Buffer, Length := 2048);
   PayloadSize := UINT_TO_UDINT(RecordCount) * UINT_TO_UDINT(RecordSize);
   TotalSize := UINT_TO_UDINT(NH_API_HEADER_SIZE) + PayloadSize;
   FrameRevision := NhApiNextRevision(Current := NhApiInfo.TxPublishedRevision);
   NhApiWriteU32(Buffer := Buffer, Offset := 0, Value := DWORD_TO_UDINT(NH_API_MAGIC));
   NhApiWriteU16(Buffer := Buffer, Offset := 4, Value := NH_API_PROTOCOL_VERSION);
   NhApiWriteU16(Buffer := Buffer, Offset := 6, Value := NH_API_HEADER_SIZE);
   NhApiWriteU16(Buffer := Buffer, Offset := 8, Value := MessageType);
   NhApiWriteU16(Buffer := Buffer, Offset := 10, Value := SchemaId);
   NhApiWriteU16(Buffer := Buffer, Offset := 12, Value := NH_API_SCHEMA_VERSION);
   NhApiWriteU16(Buffer := Buffer, Offset := 14, Value := 0);
   NhApiWriteU32(Buffer := Buffer, Offset := 16, Value := 0);
   NhApiWriteU32(Buffer := Buffer, Offset := 20, Value := RequestId);
   NhApiWriteU32(Buffer := Buffer, Offset := 24, Value := FrameRevision);
   NhApiWriteU32(Buffer := Buffer, Offset := 28, Value := FromRevision);
   NhApiWriteU32(Buffer := Buffer, Offset := 32, Value := ToRevision);
   NhApiWriteU16(Buffer := Buffer, Offset := 36, Value := RecordCount);
   NhApiWriteU16(Buffer := Buffer, Offset := 38, Value := RecordSize);
   NhApiWriteU16(Buffer := Buffer, Offset := 40, Value := PartIndex);
   NhApiWriteU16(Buffer := Buffer, Offset := 42, Value := PartCount);
   NhApiWriteU32(Buffer := Buffer, Offset := 44, Value := PayloadSize);
   NhApiWriteU32(Buffer := Buffer, Offset := 48, Value := TargetClientId);
   NhApiWriteU16(Buffer := Buffer, Offset := 52, Value := USINT_TO_UINT(NH_API_RESULT_OK));
   NhApiWriteU16(Buffer := Buffer, Offset := 54, Value := 0);
   NhApiWriteU32(Buffer := Buffer, Offset := 56, Value := TotalSize);
   NhApiWriteU32(Buffer := Buffer, Offset := 60, Value := 0);
   NhApiInfo.TxByteLength := UDINT_TO_UINT(TotalSize);
   NhApiBeginFrame := TRUE;
END_FUNCTION

FUNCTION NhApiPublishFrame : BOOL
   // Adds CRC and atomically publishes the prepared TX frame. SK: Doplni CRC a atomicky publikuje pripraveny TX ramec.
   VAR
      Buffer : PTR_TO BYTE; // Byte view of the TX DWORD array. SK: Byte pohlad na TX DWORD pole.
      Crc : DWORD;          // CRC32 of the complete valid frame. SK: CRC32 celeho platneho ramca.
   END_VAR
   Buffer := ADR(NhApiTxBuffer);
   Crc := NhApiFrameCrc32(Buffer := Buffer, Length := NhApiInfo.TxByteLength);
   NhApiWriteU32(Buffer := Buffer, Offset := 60, Value := DWORD_TO_UDINT(Crc));
   NhApiInfo.TxPublishedRevision := NhApiReadU32(Buffer := Buffer, Offset := 24);
   NhApiInfo.TxRequiredAckMask := NhApiInfo.ActiveClientMask;
   NhApiInfo.TxAckMask := 0;
   NhApiInfo.TxState := NH_API_TX_READY;
   NhApiPublishFrame := TRUE;
END_FUNCTION

FUNCTION NhApiStartSnapshot : BOOL
   // Freezes current room data and starts the snapshot sequence. SK: Zmrazi aktualne room data a spusti sekvenciu snapshotu.
   VAR_INPUT
      TargetClientId : UDINT; // Zero for a WebMaker broadcast. SK: Nula pre WebMaker broadcast.
      RequestId : UDINT;      // Request identifier. SK: Identifikator poziadavky.
   END_VAR
   VAR
      Index : USINT;          // Source room slot. SK: Zdrojovy room slot.
   END_VAR
   NhApiStartSnapshot := FALSE;
   IF NhSnapshotActive OR (NhPendingKind <> 0) OR (NhApiInfo.TxState <> NH_API_TX_IDLE) THEN
      RETURN;
   END_IF;
   NhSnapshotCount := 0;
   FOR Index := 1 TO NH_API_MAX_ROOMS DO
      IF NhRoomsConfig[Index].Used THEN
         NhSnapshotCount := NhSnapshotCount + 1;
         NhSnapshotConfig[NhSnapshotCount] := NhRoomsConfig[Index];
         NhSnapshotState[NhSnapshotCount] := NhRoomsState[Index];
      END_IF;
   END_FOR;
   NhSnapshotActive := TRUE;
   NhSnapshotTargetClientId := TargetClientId;
   NhSnapshotRequestId := RequestId;
   NhSnapshotStage := 1;
   NhSnapshotNext := 1;
   NhSnapshotPart := 1;
   NhSnapshotParts := (NhSnapshotCount + NH_API_CONFIG_PER_FRAME - 1) / NH_API_CONFIG_PER_FRAME;
   IF NhSnapshotParts = 0 THEN
      NhSnapshotParts := 1;
   END_IF;
   NhApiStartSnapshot := TRUE;
END_FUNCTION

FUNCTION NhApiPublishSnapshotPart : BOOL
   // Builds and publishes one part of the active snapshot. SK: Vytvori a publikuje jednu cast rozpracovaneho snapshotu.
   VAR
      Buffer : PTR_TO BYTE; // Byte view of the TX buffer. SK: Byte pohlad na TX buffer.
      Count : USINT;        // Number of records in this part. SK: Pocet zaznamov tejto casti.
      Index : USINT;        // Local record index. SK: Lokalny index zaznamu.
      Source : USINT;       // Index in the frozen snapshot. SK: Index v zmrazenom snapshote.
      Offset : UINT;        // Record byte offset. SK: Byte offset zaznamu.
   END_VAR
   NhApiPublishSnapshotPart := FALSE;
   IF NOT NhSnapshotActive OR (NhApiInfo.TxState <> NH_API_TX_IDLE) THEN
      RETURN;
   END_IF;
   Buffer := ADR(NhApiTxBuffer);
   IF NhSnapshotStage = 1 THEN
      Count := NH_API_CONFIG_PER_FRAME;
      IF (NhSnapshotNext + Count - 1) > NhSnapshotCount THEN
         Count := NhSnapshotCount - NhSnapshotNext + 1;
      END_IF;
      NhApiBeginFrame(MessageType := NH_API_MSG_CONFIG_SNAPSHOT, SchemaId := NH_API_SCHEMA_ROOM_CONFIG,
         TargetClientId := NhSnapshotTargetClientId, RequestId := NhSnapshotRequestId,
         FromRevision := 0, ToRevision := NhApiInfo.ConfigRevision, RecordCount := USINT_TO_UINT(Count),
         RecordSize := NH_API_CONFIG_RECORD_SIZE, PartIndex := USINT_TO_UINT(NhSnapshotPart),
         PartCount := USINT_TO_UINT(NhSnapshotParts));
      FOR Index := 0 TO Count - 1 DO
         Source := NhSnapshotNext + Index;
         Offset := NH_API_HEADER_SIZE + USINT_TO_UINT(Index) * NH_API_CONFIG_RECORD_SIZE;
         NhApiWriteConfigRecord(Buffer := Buffer, Offset := Offset, Record := NhSnapshotConfig[Source]);
      END_FOR;
      NhSnapshotNext := NhSnapshotNext + Count;
      NhSnapshotPart := NhSnapshotPart + 1;
      IF NhSnapshotNext > NhSnapshotCount THEN
         NhSnapshotStage := 2;
         NhSnapshotNext := 1;
         NhSnapshotPart := 1;
         NhSnapshotParts := (NhSnapshotCount + NH_API_STATE_PER_FRAME - 1) / NH_API_STATE_PER_FRAME;
         IF NhSnapshotParts = 0 THEN NhSnapshotParts := 1; END_IF;
      END_IF;
   ELSIF NhSnapshotStage = 2 THEN
      Count := NH_API_STATE_PER_FRAME;
      IF (NhSnapshotNext + Count - 1) > NhSnapshotCount THEN
         Count := NhSnapshotCount - NhSnapshotNext + 1;
      END_IF;
      NhApiBeginFrame(MessageType := NH_API_MSG_STATE_SNAPSHOT, SchemaId := NH_API_SCHEMA_ROOM_STATE,
         TargetClientId := NhSnapshotTargetClientId, RequestId := NhSnapshotRequestId,
         FromRevision := 0, ToRevision := NhApiInfo.StateRevision, RecordCount := USINT_TO_UINT(Count),
         RecordSize := NH_API_STATE_RECORD_SIZE, PartIndex := USINT_TO_UINT(NhSnapshotPart),
         PartCount := USINT_TO_UINT(NhSnapshotParts));
      FOR Index := 0 TO Count - 1 DO
         Source := NhSnapshotNext + Index;
         Offset := NH_API_HEADER_SIZE + USINT_TO_UINT(Index) * NH_API_STATE_RECORD_SIZE;
         NhApiWriteStateRecord(Buffer := Buffer, Offset := Offset, Record := NhSnapshotState[Source]);
      END_FOR;
      NhSnapshotNext := NhSnapshotNext + Count;
      NhSnapshotPart := NhSnapshotPart + 1;
      IF NhSnapshotNext > NhSnapshotCount THEN
         NhSnapshotStage := 3;
      END_IF;
   ELSIF NhSnapshotStage = 3 THEN
      NhApiBeginFrame(MessageType := NH_API_MSG_SNAPSHOT_DONE, SchemaId := NH_API_SCHEMA_NONE,
         TargetClientId := NhSnapshotTargetClientId, RequestId := NhSnapshotRequestId,
         FromRevision := NhApiInfo.ConfigRevision, ToRevision := NhApiInfo.StateRevision,
         RecordCount := 0, RecordSize := 0, PartIndex := 1, PartCount := 1);
      NhSnapshotStage := 4;
   ELSE
      NhSnapshotActive := FALSE;
      RETURN;
   END_IF;
   NhApiPublishFrame();
   NhApiPublishSnapshotPart := TRUE;
END_FUNCTION

FUNCTION NhApiCaptureConfigDiff : BOOL
   // Captures configuration changes into a frozen pending diff. SK: Zachyti konfiguracne zmeny a zmrazi ich do pending diffu.
   VAR
      Index : USINT; // Room slot. SK: Room slot.
   END_VAR
   NhApiCaptureConfigDiff := FALSE;
   NhPendingCount := 0;
   FOR Index := 1 TO NH_API_MAX_ROOMS DO
      IF NOT NhApiConfigEqual(A := NhRoomsConfig[Index], B := NhConfigShadow[Index]) THEN
         NhPendingCount := NhPendingCount + 1;
         IF NhRoomsConfig[Index].Used THEN
            NhPendingOperation[NhPendingCount] := NH_API_CHANGE_UPSERT;
            NhPendingRoomId[NhPendingCount] := NhRoomsConfig[Index].RoomId;
            NhPendingConfig[NhPendingCount] := NhRoomsConfig[Index];
         ELSE
            NhPendingOperation[NhPendingCount] := NH_API_CHANGE_DELETE;
            NhPendingRoomId[NhPendingCount] := NhConfigShadow[Index].RoomId;
            NhPendingConfig[NhPendingCount] := NhRoomsConfig[Index];
         END_IF;
         NhConfigShadow[Index] := NhRoomsConfig[Index];
      END_IF;
   END_FOR;
   IF NhPendingCount > 0 THEN
      NhPendingKind := NH_API_MSG_CONFIG_DIFF;
      NhPendingFromRevision := NhApiInfo.ConfigRevision;
      NhApiInfo.ConfigRevision := NhApiNextRevision(Current := NhApiInfo.ConfigRevision);
      NhPendingToRevision := NhApiInfo.ConfigRevision;
      NhPendingNext := 1;
      NhPendingPart := 1;
      NhPendingParts := (NhPendingCount + NH_API_CONFIG_DIFF_PER_FRAME - 1) / NH_API_CONFIG_DIFF_PER_FRAME;
      NhApiCaptureConfigDiff := TRUE;
   END_IF;
END_FUNCTION

FUNCTION NhApiCaptureStateDiff : BOOL
   // Captures state changes into a frozen pending diff. SK: Zachyti stavove zmeny a zmrazi ich do pending diffu.
   VAR
      Index : USINT; // Room slot. SK: Room slot.
   END_VAR
   NhApiCaptureStateDiff := FALSE;
   NhPendingCount := 0;
   FOR Index := 1 TO NH_API_MAX_ROOMS DO
      IF NOT NhApiStateEqual(A := NhRoomsState[Index], B := NhStateShadow[Index]) THEN
         NhPendingCount := NhPendingCount + 1;
         IF NhRoomsConfig[Index].Used THEN
            NhPendingOperation[NhPendingCount] := NH_API_CHANGE_UPSERT;
            NhPendingRoomId[NhPendingCount] := NhRoomsState[Index].RoomId;
            NhPendingState[NhPendingCount] := NhRoomsState[Index];
         ELSE
            NhPendingOperation[NhPendingCount] := NH_API_CHANGE_DELETE;
            NhPendingRoomId[NhPendingCount] := NhStateShadow[Index].RoomId;
            NhPendingState[NhPendingCount] := NhRoomsState[Index];
         END_IF;
         NhStateShadow[Index] := NhRoomsState[Index];
      END_IF;
   END_FOR;
   IF NhPendingCount > 0 THEN
      NhPendingKind := NH_API_MSG_STATE_DIFF;
      NhPendingFromRevision := NhApiInfo.StateRevision;
      NhApiInfo.StateRevision := NhApiNextRevision(Current := NhApiInfo.StateRevision);
      NhPendingToRevision := NhApiInfo.StateRevision;
      NhPendingNext := 1;
      NhPendingPart := 1;
      NhPendingParts := (NhPendingCount + NH_API_STATE_DIFF_PER_FRAME - 1) / NH_API_STATE_DIFF_PER_FRAME;
      NhApiCaptureStateDiff := TRUE;
   END_IF;
END_FUNCTION

FUNCTION NhApiPublishPendingDiff : BOOL
   // Builds and publishes one part of the frozen diff. SK: Vytvori a publikuje jednu cast zmrazeneho diffu.
   // The frame contains only one schema and one diff section. SK: Ramec obsahuje iba jednu schemu a jednu diff sekciu.
   VAR
      Buffer : PTR_TO BYTE; // Byte view of the TX buffer. SK: Byte pohlad na TX buffer.
      Count : USINT;        // Number of changes in this part. SK: Pocet zmien tejto casti.
      Index : USINT;        // Local change index. SK: Lokalny index zmeny.
      Source : USINT;       // Frozen change index. SK: Index zmrazenej zmeny.
      Offset : UINT;        // Change byte offset. SK: Byte offset zmeny.
   END_VAR
   NhApiPublishPendingDiff := FALSE;
   IF (NhPendingKind = 0) OR (NhApiInfo.TxState <> NH_API_TX_IDLE) THEN RETURN; END_IF;
   Buffer := ADR(NhApiTxBuffer);
   IF NhPendingKind = NH_API_MSG_CONFIG_DIFF THEN
      Count := NH_API_CONFIG_DIFF_PER_FRAME;
      IF (NhPendingNext + Count - 1) > NhPendingCount THEN Count := NhPendingCount - NhPendingNext + 1; END_IF;
      NhApiBeginFrame(MessageType := NH_API_MSG_CONFIG_DIFF, SchemaId := NH_API_SCHEMA_ROOM_CONFIG,
         TargetClientId := 0, RequestId := 0, FromRevision := NhPendingFromRevision,
         ToRevision := NhPendingToRevision, RecordCount := USINT_TO_UINT(Count),
         RecordSize := NH_API_CONFIG_DIFF_SIZE, PartIndex := USINT_TO_UINT(NhPendingPart),
         PartCount := USINT_TO_UINT(NhPendingParts));
      FOR Index := 0 TO Count - 1 DO
         Source := NhPendingNext + Index;
         Offset := NH_API_HEADER_SIZE + USINT_TO_UINT(Index) * NH_API_CONFIG_DIFF_SIZE;
         NhApiWriteByte(Buffer := Buffer, Offset := Offset, Value := USINT_TO_BYTE(NhPendingOperation[Source]));
         NhApiWriteU32(Buffer := Buffer, Offset := Offset + 1, Value := NhPendingRoomId[Source]);
         NhApiWriteConfigRecord(Buffer := Buffer, Offset := Offset + 5, Record := NhPendingConfig[Source]);
      END_FOR;
   ELSE
      Count := NH_API_STATE_DIFF_PER_FRAME;
      IF (NhPendingNext + Count - 1) > NhPendingCount THEN Count := NhPendingCount - NhPendingNext + 1; END_IF;
      NhApiBeginFrame(MessageType := NH_API_MSG_STATE_DIFF, SchemaId := NH_API_SCHEMA_ROOM_STATE,
         TargetClientId := 0, RequestId := 0, FromRevision := NhPendingFromRevision,
         ToRevision := NhPendingToRevision, RecordCount := USINT_TO_UINT(Count),
         RecordSize := NH_API_STATE_DIFF_SIZE, PartIndex := USINT_TO_UINT(NhPendingPart),
         PartCount := USINT_TO_UINT(NhPendingParts));
      FOR Index := 0 TO Count - 1 DO
         Source := NhPendingNext + Index;
         Offset := NH_API_HEADER_SIZE + USINT_TO_UINT(Index) * NH_API_STATE_DIFF_SIZE;
         NhApiWriteByte(Buffer := Buffer, Offset := Offset, Value := USINT_TO_BYTE(NhPendingOperation[Source]));
         NhApiWriteU32(Buffer := Buffer, Offset := Offset + 1, Value := NhPendingRoomId[Source]);
         NhApiWriteStateRecord(Buffer := Buffer, Offset := Offset + 5, Record := NhPendingState[Source]);
      END_FOR;
   END_IF;
   NhPendingNext := NhPendingNext + Count;
   NhPendingPart := NhPendingPart + 1;
   IF NhPendingNext > NhPendingCount THEN NhPendingKind := 0; END_IF;
   NhApiPublishFrame();
   NhApiPublishPendingDiff := TRUE;
END_FUNCTION

FUNCTION NhApiApplyAdd : USINT
   // Adds a new room to the first free slot. SK: Prida novu miestnost do prveho volneho slotu.
   VAR_INPUT
      Record : NH_ROOM_CONFIG; // New configuration. SK: Nova konfiguracia.
   END_VAR
   VAR
      Slot : USINT;              // Free internal slot. SK: Volny interny slot.
   END_VAR
   IF (Record.RoomId = 0) OR (LEN(Record.Name) = 0) THEN NhApiApplyAdd := NH_API_RESULT_INVALID; RETURN; END_IF;
   IF NhApiFindRoom(RoomId := Record.RoomId) <> 0 THEN NhApiApplyAdd := NH_API_RESULT_ALREADY_EXISTS; RETURN; END_IF;
   Slot := NhApiFindFreeRoom();
   IF Slot = 0 THEN NhApiApplyAdd := NH_API_RESULT_NO_FREE_SLOT; RETURN; END_IF;
   NhRoomsConfig[Slot] := Record;
   NhRoomsConfig[Slot].Used := TRUE;
   IF NhRoomsConfig[Slot].IconId = 0 THEN NhRoomsConfig[Slot].IconId := 16; END_IF;
   IF NhRoomsConfig[Slot].SortDefault = 0 THEN NhRoomsConfig[Slot].SortDefault := USINT_TO_UINT(Slot); END_IF;
   NhRoomsState[Slot].RoomId := Record.RoomId;
   NhRoomsState[Slot].Temperature := 20.0;
   NhRoomsState[Slot].Humidity := 40.0;
   NhRoomsState[Slot].Presence := FALSE;
   NhRoomsState[Slot].DayPhase := 140;
   NhRoomsState[Slot].CategoryMask := 0;
   NhRoomsState[Slot].AlarmLevel := 0;
   NhRoomsState[Slot].Online := TRUE;
   NhRoomsState[Slot].Twilight := FALSE;
   NhApiApplyAdd := NH_API_RESULT_OK;
END_FUNCTION

FUNCTION NhApiApplyDelete : USINT
   // Deletes a room by its stable ID. SK: Odstrani miestnost podla jej stabilneho ID.
   VAR_INPUT
      RoomId : UDINT;             // ID of the room to delete. SK: ID mazanej miestnosti.
   END_VAR
   VAR
      Slot : USINT;               // Located internal slot. SK: Najdeny interny slot.
   END_VAR
   Slot := NhApiFindRoom(RoomId := RoomId);
   IF Slot = 0 THEN NhApiApplyDelete := NH_API_RESULT_NOT_FOUND; RETURN; END_IF;
   NhApiClearRoom(Index := Slot);
   NhApiApplyDelete := NH_API_RESULT_OK;
END_FUNCTION

FUNCTION NhApiApplyConfig : USINT
   // Replaces the configuration of an existing room. SK: Nahradi konfiguraciu existujucej miestnosti.
   VAR_INPUT
      Record : NH_ROOM_CONFIG;  // Complete new configuration. SK: Uplna nova konfiguracia.
   END_VAR
   VAR
      Slot : USINT;               // Located internal slot. SK: Najdeny interny slot.
   END_VAR
   Slot := NhApiFindRoom(RoomId := Record.RoomId);
   IF Slot = 0 THEN NhApiApplyConfig := NH_API_RESULT_NOT_FOUND; RETURN; END_IF;
   IF LEN(Record.Name) = 0 THEN NhApiApplyConfig := NH_API_RESULT_INVALID; RETURN; END_IF;
   NhRoomsConfig[Slot] := Record;
   NhRoomsConfig[Slot].Used := TRUE;
   NhApiApplyConfig := NH_API_RESULT_OK;
END_FUNCTION

FUNCTION NhApiApplyState : USINT
   // Replaces the dynamic state of an existing room. SK: Nahradi dynamicky stav existujucej miestnosti.
   VAR_INPUT
      Record : NH_ROOM_STATE;   // Complete new dynamic state. SK: Uplny novy dynamicky stav.
   END_VAR
   VAR
      Slot : USINT;               // Located internal slot. SK: Najdeny interny slot.
   END_VAR
   Slot := NhApiFindRoom(RoomId := Record.RoomId);
   IF Slot = 0 THEN NhApiApplyState := NH_API_RESULT_NOT_FOUND; RETURN; END_IF;
   IF (Record.Temperature < -50.0) OR (Record.Temperature > 100.0) OR
      (Record.Humidity < 0.0) OR (Record.Humidity > 100.0) OR (Record.AlarmLevel > 2) THEN
      NhApiApplyState := NH_API_RESULT_INVALID; RETURN;
   END_IF;
   NhRoomsState[Slot] := Record;
   NhApiApplyState := NH_API_RESULT_OK;
END_FUNCTION

FUNCTION NhApiApplyCopy : USINT
   // Creates a new room by copying an existing one. SK: Vytvori novu miestnost skopirovanim existujucej.
   VAR_INPUT
      SourceRoomId : UDINT;       // Source room ID. SK: ID zdrojovej miestnosti.
      Target       : NH_ROOM_CONFIG; // Target ID and optional new config fields. SK: Cielove ID a volitelne nove config polia.
   END_VAR
   VAR
      SourceSlot : USINT;         // Source internal slot. SK: Zdrojovy interny slot.
      TargetSlot : USINT;         // Target free slot. SK: Cielovy volny slot.
   END_VAR
   SourceSlot := NhApiFindRoom(RoomId := SourceRoomId);
   IF SourceSlot = 0 THEN NhApiApplyCopy := NH_API_RESULT_NOT_FOUND; RETURN; END_IF;
   IF (Target.RoomId = 0) OR (NhApiFindRoom(RoomId := Target.RoomId) <> 0) THEN NhApiApplyCopy := NH_API_RESULT_ALREADY_EXISTS; RETURN; END_IF;
   TargetSlot := NhApiFindFreeRoom();
   IF TargetSlot = 0 THEN NhApiApplyCopy := NH_API_RESULT_NO_FREE_SLOT; RETURN; END_IF;
   NhRoomsConfig[TargetSlot] := NhRoomsConfig[SourceSlot];
   NhRoomsConfig[TargetSlot].RoomId := Target.RoomId;
   NhRoomsConfig[TargetSlot].SortDefault := USINT_TO_UINT(TargetSlot);
   IF LEN(Target.Name) > 0 THEN NhRoomsConfig[TargetSlot].Name := Target.Name; END_IF;
   IF LEN(Target.ProjectName) > 0 THEN NhRoomsConfig[TargetSlot].ProjectName := Target.ProjectName; END_IF;
   IF Target.IconId > 0 THEN NhRoomsConfig[TargetSlot].IconId := Target.IconId; END_IF;
   NhRoomsState[TargetSlot] := NhRoomsState[SourceSlot];
   NhRoomsState[TargetSlot].RoomId := Target.RoomId;
   NhApiApplyCopy := NH_API_RESULT_OK;
END_FUNCTION

FUNCTION NhApiProcessClients : BOOL
   // Maintains the client registry, timeouts, and TX acknowledgements. SK: Udrzuje registry klientov, timeouty a potvrdenia TX ramca.
   VAR
      Index : USINT;              // Client slot. SK: Klientsky slot.
      NowMs : UDINT;              // System millisecond time. SK: Systemovy milisekundovy cas.
      BitMask : BYTE;             // Bit belonging to the client. SK: Bit prisluchajuci klientovi.
      Activity : BOOL;            // Client changed heartbeat, ACK or RX. SK: Klient zmenil heartbeat, ACK alebo RX.
   END_VAR
   NowMs := NhApiSystemTimeMs();
   NhApiInfo.ActiveClientMask := 0;
   NhApiInfo.TxAckMask := 0;
   FOR Index := 0 TO 3 DO
      BitMask := SHL(BYTE#1, USINT_TO_UINT(Index));
      IF NhApiClients[Index].State = NH_API_CLIENT_FREE THEN
         IF NhApiClients[Index].RequestedClientId <> 0 THEN
            NhApiClients[Index].AssignedClientId := NhApiClients[Index].RequestedClientId;
            NhApiClients[Index].State := NH_API_CLIENT_ACTIVE;
            NhClientLastHeartbeat[Index] := NhApiClients[Index].HeartbeatCounter;
            NhClientLastAck[Index] := NhApiClients[Index].AckTxRevision;
            NhClientLastRx[Index] := NhApiClients[Index].RxPublishedRevision;
            NhClientLastActivityMs[Index] := NowMs;
         END_IF;
      ELSE
         Activity := (NhApiClients[Index].HeartbeatCounter <> NhClientLastHeartbeat[Index]) OR
            (NhApiClients[Index].AckTxRevision <> NhClientLastAck[Index]) OR
            (NhApiClients[Index].RxPublishedRevision <> NhClientLastRx[Index]);
         IF Activity THEN
            NhClientLastHeartbeat[Index] := NhApiClients[Index].HeartbeatCounter;
            NhClientLastAck[Index] := NhApiClients[Index].AckTxRevision;
            NhClientLastActivityMs[Index] := NowMs;
         END_IF;
         IF (NhApiClients[Index].RequestedClientId = 0) OR
            ((NowMs - NhClientLastActivityMs[Index]) > NH_API_CLIENT_TIMEOUT_MS) THEN
            NhApiClients[Index].RequestedClientId := 0;
            NhApiClients[Index].AssignedClientId := 0;
            NhApiClients[Index].State := NH_API_CLIENT_FREE;
            NhApiClients[Index].ResultCode := NH_API_RESULT_NONE;
         END_IF;
      END_IF;
      IF NhApiClients[Index].State = NH_API_CLIENT_ACTIVE THEN
         NhApiInfo.ActiveClientMask := NhApiInfo.ActiveClientMask OR BitMask;
         IF NhApiClients[Index].AckTxRevision = NhApiInfo.TxPublishedRevision THEN
            NhApiInfo.TxAckMask := NhApiInfo.TxAckMask OR BitMask;
         END_IF;
      END_IF;
   END_FOR;
   IF NhApiInfo.TxState = NH_API_TX_READY THEN
      NhApiInfo.TxRequiredAckMask := NhApiInfo.TxRequiredAckMask AND NhApiInfo.ActiveClientMask;
      IF (NhApiInfo.TxAckMask AND NhApiInfo.TxRequiredAckMask) = NhApiInfo.TxRequiredAckMask THEN
         NhApiInfo.TxState := NH_API_TX_IDLE;
         NhApiInfo.TxRequiredAckMask := 0;
      END_IF;
   END_IF;
   NhApiProcessClients := TRUE;
END_FUNCTION

FUNCTION NhApiProcessOneRx : BOOL
   // Validates and processes at most one new client RX request. SK: Overi a spracuje najviac jednu novu klientsku RX poziadavku.
   VAR
      Index : USINT;              // Client slot. SK: Klientsky slot.
      BaseWord : UINT;            // First DWORD of the client RX segment. SK: Prvy DWORD klientovho RX segmentu.
      Buffer : PTR_TO BYTE;       // Byte view of the RX segment. SK: Byte pohlad na RX segment.
      Length : UINT;              // Declared RX frame size. SK: Deklarovana velkost RX ramca.
      MessageType : UINT;         // RX request type. SK: Typ RX poziadavky.
      ClientId : UDINT;           // ClientId from the header. SK: ClientId z hlavicky.
      RequestId : UDINT;          // RequestId from the header. SK: RequestId z hlavicky.
      ExpectedCrc : DWORD;        // CRC written by the client. SK: CRC zapisane klientom.
      ActualCrc : DWORD;          // CRC calculated by the PLC. SK: CRC vypocitane PLC.
      Result : USINT;             // Executed operation result. SK: Vysledok vykonanej operacie.
      ConfigRecord : NH_ROOM_CONFIG; // Decoded config record. SK: Dekodovany config zaznam.
      StateRecord : NH_ROOM_STATE;   // Decoded state record. SK: Dekodovany state zaznam.
      SourceRoomId : UDINT;       // Source ID for copy command. SK: Zdrojove ID prikazu copy.
   END_VAR
   NhApiProcessOneRx := FALSE;
   IF (NhApiInfo.TxState <> NH_API_TX_IDLE) OR NhSnapshotActive OR (NhPendingKind <> 0) THEN RETURN; END_IF;
   FOR Index := 0 TO 3 DO
      IF (NhApiClients[Index].State = NH_API_CLIENT_ACTIVE) AND
         (NhApiClients[Index].RxPublishedRevision <> NhClientLastRx[Index]) THEN
         BaseWord := USINT_TO_UINT(Index) * NH_API_RX_WORDS_PER_CLIENT;
         Buffer := ADR(NhApiRxBuffer[BaseWord]);
         Length := NhApiClients[Index].RxByteLength;
         Result := NH_API_RESULT_BAD_FRAME;
         RequestId := 0;
         IF (Length >= NH_API_HEADER_SIZE) AND (Length <= 256) AND
            (NhApiReadU32(Buffer := Buffer, Offset := 0) = DWORD_TO_UDINT(NH_API_MAGIC)) AND
            (NhApiReadU16(Buffer := Buffer, Offset := 4) = NH_API_PROTOCOL_VERSION) AND
            (NhApiReadU16(Buffer := Buffer, Offset := 6) = NH_API_HEADER_SIZE) AND
            (NhApiReadU32(Buffer := Buffer, Offset := 24) = NhApiClients[Index].RxPublishedRevision) AND
            ((NhApiReadU32(Buffer := Buffer, Offset := 44) + UINT_TO_UDINT(NH_API_HEADER_SIZE)) = UINT_TO_UDINT(Length)) AND
            (NhApiReadU32(Buffer := Buffer, Offset := 56) = UINT_TO_UDINT(Length)) THEN
            ExpectedCrc := UDINT_TO_DWORD(NhApiReadU32(Buffer := Buffer, Offset := 60));
            ActualCrc := NhApiFrameCrc32(Buffer := Buffer, Length := Length);
            ClientId := NhApiReadU32(Buffer := Buffer, Offset := 16);
            RequestId := NhApiReadU32(Buffer := Buffer, Offset := 20);
            MessageType := NhApiReadU16(Buffer := Buffer, Offset := 8);
            IF (ExpectedCrc = ActualCrc) AND (ClientId = NhApiClients[Index].AssignedClientId) AND (RequestId <> 0) THEN
               IF RequestId = NhApiClients[Index].LastRequestId THEN
                  Result := NhApiClients[Index].ResultCode;
               ELSE
                  CASE MessageType OF
                     NH_API_MSG_SNAPSHOT_REQUEST:
                        IF NhApiStartSnapshot(TargetClientId := ClientId, RequestId := RequestId) THEN Result := NH_API_RESULT_OK; ELSE Result := NH_API_RESULT_BUSY; END_IF;
                     NH_API_MSG_ADD_ROOM:
                        NhApiReadConfigRecord(Buffer := Buffer, Offset := NH_API_HEADER_SIZE, Record := ConfigRecord);
                        Result := NhApiApplyAdd(Record := ConfigRecord);
                     NH_API_MSG_DELETE_ROOM:
                        Result := NhApiApplyDelete(RoomId := NhApiReadU32(Buffer := Buffer, Offset := NH_API_HEADER_SIZE));
                     NH_API_MSG_COPY_ROOM:
                        SourceRoomId := NhApiReadU32(Buffer := Buffer, Offset := NH_API_HEADER_SIZE);
                        NhApiReadConfigRecord(Buffer := Buffer, Offset := NH_API_HEADER_SIZE + 4, Record := ConfigRecord);
                        Result := NhApiApplyCopy(SourceRoomId := SourceRoomId, Target := ConfigRecord);
                     NH_API_MSG_SET_ROOM_CONFIG:
                        NhApiReadConfigRecord(Buffer := Buffer, Offset := NH_API_HEADER_SIZE, Record := ConfigRecord);
                        Result := NhApiApplyConfig(Record := ConfigRecord);
                     NH_API_MSG_SET_ROOM_STATE:
                        NhApiReadStateRecord(Buffer := Buffer, Offset := NH_API_HEADER_SIZE, Record := StateRecord);
                        Result := NhApiApplyState(Record := StateRecord);
                     ELSE
                        Result := NH_API_RESULT_UNSUPPORTED;
                  END_CASE;
               END_IF;
            END_IF;
         END_IF;
         NhClientLastRx[Index] := NhApiClients[Index].RxPublishedRevision;
         NhClientLastActivityMs[Index] := NhApiSystemTimeMs();
         NhApiClients[Index].LastRequestId := RequestId;
         NhApiClients[Index].ResultCode := Result;
         NhApiClients[Index].ResultConfigRevision := NhApiInfo.ConfigRevision;
         NhApiClients[Index].ResultStateRevision := NhApiInfo.StateRevision;
         NhApiProcessOneRx := TRUE;
         RETURN;
      END_IF;
   END_FOR;
END_FUNCTION

FUNCTION NhApiProcessTest : BOOL
   // Processes one test action submitted through WebMaker. SK: Spracuje jednu testovaciu akciu zadanu cez WebMaker.
   VAR
      Slot : USINT;               // Located room slot. SK: Najdeny room slot.
      Result : USINT;             // WebMaker action result. SK: Vysledok WebMaker akcie.
      ConfigRecord : NH_ROOM_CONFIG; // Constructed config record. SK: Zostaveny config zaznam.
      StateRecord : NH_ROOM_STATE;   // Constructed state record. SK: Zostaveny state zaznam.
   END_VAR
   NhApiProcessTest := FALSE;
   IF NOT NhApiTest.Execute THEN RETURN; END_IF;
   IF (NhApiInfo.TxState <> NH_API_TX_IDLE) OR NhSnapshotActive OR (NhPendingKind <> 0) THEN
      NhApiTest.Busy := TRUE;
      NhApiTest.Finished := FALSE;
      RETURN;
   END_IF;
   NhApiTest.Busy := TRUE;
   NhApiTest.Finished := FALSE;
   Result := NH_API_RESULT_UNSUPPORTED;
   IF NhApiTest.Action = NH_API_TEST_REQUEST_SNAPSHOT THEN
      IF NhApiStartSnapshot(TargetClientId := 0, RequestId := 0) THEN Result := NH_API_RESULT_OK; ELSE Result := NH_API_RESULT_BUSY; END_IF;
   ELSIF NhApiTest.Action = NH_API_TEST_DELETE_ROOM THEN
      Result := NhApiApplyDelete(RoomId := NhApiTest.RoomId);
   ELSIF NhApiTest.Action = NH_API_TEST_SET_STATE THEN
      Slot := NhApiFindRoom(RoomId := NhApiTest.RoomId);
      IF Slot = 0 THEN
         Result := NH_API_RESULT_NOT_FOUND;
      ELSE
         StateRecord := NhRoomsState[Slot];
         StateRecord.Temperature := NhApiTest.Temperature;
         StateRecord.Humidity := NhApiTest.Humidity;
         StateRecord.Presence := NhApiTest.Presence;
         StateRecord.DayPhase := NhApiTest.DayPhase;
         StateRecord.CategoryMask := NhApiTest.CategoryMask;
         StateRecord.AlarmLevel := NhApiTest.AlarmLevel;
         StateRecord.Online := NhApiTest.Online;
         StateRecord.Twilight := NhApiTest.Twilight;
         Result := NhApiApplyState(Record := StateRecord);
      END_IF;
   ELSE
      ConfigRecord.Used := TRUE;
      ConfigRecord.RoomId := NhApiTest.RoomId;
      ConfigRecord.Name := NhApiTest.Name;
      ConfigRecord.ProjectName := NhApiTest.ProjectName;
      ConfigRecord.IconId := NhApiTest.IconId;
      ConfigRecord.SortDefault := 0;
      IF NhApiTest.Action = NH_API_TEST_ADD_ROOM THEN
         Result := NhApiApplyAdd(Record := ConfigRecord);
      ELSIF NhApiTest.Action = NH_API_TEST_COPY_ROOM THEN
         Result := NhApiApplyCopy(SourceRoomId := NhApiTest.SourceRoomId, Target := ConfigRecord);
      ELSIF NhApiTest.Action = NH_API_TEST_SET_CONFIG THEN
         Slot := NhApiFindRoom(RoomId := NhApiTest.RoomId);
         IF Slot = 0 THEN
            Result := NH_API_RESULT_NOT_FOUND;
         ELSE
            ConfigRecord.SortDefault := NhRoomsConfig[Slot].SortDefault;
            Result := NhApiApplyConfig(Record := ConfigRecord);
         END_IF;
      END_IF;
   END_IF;
   NhApiTest.ResultCode := Result;
   NhApiTest.ConfigRevision := NhApiInfo.ConfigRevision;
   NhApiTest.StateRevision := NhApiInfo.StateRevision;
   NhApiTest.Execute := FALSE;
   NhApiTest.Busy := FALSE;
   NhApiTest.Finished := TRUE;
   NhApiProcessTest := TRUE;
END_FUNCTION

FUNCTION NhApiCycle : BOOL
   // Executes one cycle of the API state machine. SK: Vykona jeden cyklus stavoveho automatu API.
   VAR
      Captured : BOOL;            // A new diff was captured in this cycle. SK: V tomto cykle vznikol novy diff.
   END_VAR
   NhApiProcessClients();
   IF NhApiInfo.TxState = NH_API_TX_IDLE THEN
      IF NhSnapshotActive THEN
         NhApiPublishSnapshotPart();
      ELSIF NhPendingKind <> 0 THEN
         NhApiPublishPendingDiff();
      ELSE
         NhApiProcessOneRx();
         NhApiProcessTest();
         IF NhSnapshotActive THEN
            NhApiPublishSnapshotPart();
         ELSE
            Captured := NhApiCaptureConfigDiff();
            IF NOT Captured THEN Captured := NhApiCaptureStateDiff(); END_IF;
            IF Captured THEN NhApiPublishPendingDiff(); END_IF;
         END_IF;
      END_IF;
   END_IF;
   NhApiCycle := TRUE;
END_FUNCTION

(* ---- prgMain.ST ---- *)
PROGRAM prgMain
   // Runs initialization and one API step in every PLC cycle. SK: Spusta inicializaciu a jeden API krok v kazdom PLC cykle.
   VAR
      InitOk : BOOL; // Diagnostic result of one-time initialization. SK: Diagnosticky vysledok jednorazovej inicializacie.
      CycleOk : BOOL;// Diagnostic result of the API cycle. SK: Diagnosticky vysledok API cyklu.
   END_VAR

   // After the first cycle the function no longer overwrites authoritative data. SK: Funkcia po prvom cykle uz autoritativne data neprepisuje.
   InitOk := NhApiInitialize();
   IF InitOk THEN
      // Registry, RX, snapshot, diff and TX ACK run once per PLC cycle. SK: Registry, RX, snapshot, diff a TX ACK sa spracuju raz za PLC cyklus.
      CycleOk := NhApiCycle();
   END_IF;
END_PROGRAM
